// Tests for MONETcommon.F_WakeShakeWindow, the latched window in which the brake may stay open for the Wake&Shake (#151).
FUNCTION_BLOCK F_WakeShakeWindow_Tests EXTENDS TcUnit.FB_TestSuite
VAR
END_VAR

Sets_On_Exempt_Error();
Stays_Set_Without_Condition();
Not_Set_Stays_Not_Set();
Clear_Wins_Over_Set();
Timeout_Closes();
Park_Closes();
Covers_Not_Open_Closes();
Power_On_Closes();
Estop_Closes();
Other_Hw_Error_Closes();

// The #113 exemption opens the window.
METHOD PRIVATE Sets_On_Exempt_Error
VAR
	bWindow	: BOOL;
	sReason	: STRING(24);
END_VAR
TEST('Sets_On_Exempt_Error');
bWindow := MONETcommon.F_WakeShakeWindow(bWindow := FALSE, bSet := TRUE, bTimeout := FALSE, bParkActive := FALSE, bCoversOpen := TRUE, bPowerOnStart := FALSE, bEstop := FALSE, bOtherHwError := FALSE, sEndReason => sReason);
AssertTrue(Condition := bWindow, Message := 'window open');
AssertEquals_STRING(Expected := '', Actual := sReason, Message := 'no end reason');
TEST_FINISHED();
END_METHOD

// The exemption is gone after one scan; the window stays (the reason for the latch).
METHOD PRIVATE Stays_Set_Without_Condition
VAR
	bWindow	: BOOL;
	sReason	: STRING(24);
END_VAR
TEST('Stays_Set_Without_Condition');
bWindow := MONETcommon.F_WakeShakeWindow(bWindow := TRUE, bSet := FALSE, bTimeout := FALSE, bParkActive := FALSE, bCoversOpen := TRUE, bPowerOnStart := FALSE, bEstop := FALSE, bOtherHwError := FALSE, sEndReason => sReason);
AssertTrue(Condition := bWindow, Message := 'window stays open');
TEST_FINISHED();
END_METHOD

// No exemption, no window.
METHOD PRIVATE Not_Set_Stays_Not_Set
VAR
	bWindow	: BOOL;
	sReason	: STRING(24);
END_VAR
TEST('Not_Set_Stays_Not_Set');
bWindow := MONETcommon.F_WakeShakeWindow(bWindow := FALSE, bSet := FALSE, bTimeout := FALSE, bParkActive := FALSE, bCoversOpen := TRUE, bPowerOnStart := FALSE, bEstop := FALSE, bOtherHwError := FALSE, sEndReason => sReason);
AssertFalse(Condition := bWindow, Message := 'no window');
TEST_FINISHED();
END_METHOD

// Set and cleared in the same scan: not open, and no end reason (it never was open).
METHOD PRIVATE Clear_Wins_Over_Set
VAR
	bWindow	: BOOL;
	sReason	: STRING(24);
END_VAR
TEST('Clear_Wins_Over_Set');
bWindow := MONETcommon.F_WakeShakeWindow(bWindow := FALSE, bSet := TRUE, bTimeout := FALSE, bParkActive := FALSE, bCoversOpen := TRUE, bPowerOnStart := FALSE, bEstop := TRUE, bOtherHwError := FALSE, sEndReason => sReason);
AssertFalse(Condition := bWindow, Message := 'closed');
AssertEquals_STRING(Expected := '', Actual := sReason, Message := 'no reason');
TEST_FINISHED();
END_METHOD

// Window timer elapsed.
METHOD PRIVATE Timeout_Closes
VAR
	bWindow	: BOOL;
	sReason	: STRING(24);
END_VAR
TEST('Timeout_Closes');
bWindow := MONETcommon.F_WakeShakeWindow(bWindow := TRUE, bSet := FALSE, bTimeout := TRUE, bParkActive := FALSE, bCoversOpen := TRUE, bPowerOnStart := FALSE, bEstop := FALSE, bOtherHwError := FALSE, sEndReason => sReason);
AssertFalse(Condition := bWindow, Message := 'window closed');
AssertEquals_STRING(Expected := 'timeout', Actual := sReason, Message := 'reason');
TEST_FINISHED();
END_METHOD

// A park is requested, running or done.
METHOD PRIVATE Park_Closes
VAR
	bWindow	: BOOL;
	sReason	: STRING(24);
END_VAR
TEST('Park_Closes');
bWindow := MONETcommon.F_WakeShakeWindow(bWindow := TRUE, bSet := FALSE, bTimeout := FALSE, bParkActive := TRUE, bCoversOpen := TRUE, bPowerOnStart := FALSE, bEstop := FALSE, bOtherHwError := FALSE, sEndReason => sReason);
AssertFalse(Condition := bWindow, Message := 'window closed');
AssertEquals_STRING(Expected := 'park', Actual := sReason, Message := 'reason');
TEST_FINISHED();
END_METHOD

// The covers are not open any more.
METHOD PRIVATE Covers_Not_Open_Closes
VAR
	bWindow	: BOOL;
	sReason	: STRING(24);
END_VAR
TEST('Covers_Not_Open_Closes');
bWindow := MONETcommon.F_WakeShakeWindow(bWindow := TRUE, bSet := FALSE, bTimeout := FALSE, bParkActive := FALSE, bCoversOpen := FALSE, bPowerOnStart := FALSE, bEstop := FALSE, bOtherHwError := FALSE, sEndReason => sReason);
AssertFalse(Condition := bWindow, Message := 'window closed');
AssertEquals_STRING(Expected := 'covers not open', Actual := sReason, Message := 'reason');
TEST_FINISHED();
END_METHOD

// A new power-on enables the elevation.
METHOD PRIVATE Power_On_Closes
VAR
	bWindow	: BOOL;
	sReason	: STRING(24);
END_VAR
TEST('Power_On_Closes');
bWindow := MONETcommon.F_WakeShakeWindow(bWindow := TRUE, bSet := FALSE, bTimeout := FALSE, bParkActive := FALSE, bCoversOpen := TRUE, bPowerOnStart := TRUE, bEstop := FALSE, bOtherHwError := FALSE, sEndReason => sReason);
AssertFalse(Condition := bWindow, Message := 'window closed');
AssertEquals_STRING(Expected := 'power-on', Actual := sReason, Message := 'reason');
TEST_FINISHED();
END_METHOD

// E-stop.
METHOD PRIVATE Estop_Closes
VAR
	bWindow	: BOOL;
	sReason	: STRING(24);
END_VAR
TEST('Estop_Closes');
bWindow := MONETcommon.F_WakeShakeWindow(bWindow := TRUE, bSet := FALSE, bTimeout := FALSE, bParkActive := FALSE, bCoversOpen := TRUE, bPowerOnStart := FALSE, bEstop := TRUE, bOtherHwError := FALSE, sEndReason => sReason);
AssertFalse(Condition := bWindow, Message := 'window closed');
AssertEquals_STRING(Expected := 'E-stop', Actual := sReason, Message := 'reason');
TEST_FINISHED();
END_METHOD

// Focus or derotator error.
METHOD PRIVATE Other_Hw_Error_Closes
VAR
	bWindow	: BOOL;
	sReason	: STRING(24);
END_VAR
TEST('Other_Hw_Error_Closes');
bWindow := MONETcommon.F_WakeShakeWindow(bWindow := TRUE, bSet := FALSE, bTimeout := FALSE, bParkActive := FALSE, bCoversOpen := TRUE, bPowerOnStart := FALSE, bEstop := FALSE, bOtherHwError := TRUE, sEndReason => sReason);
AssertFalse(Condition := bWindow, Message := 'window closed');
AssertEquals_STRING(Expected := 'focus/derotator error', Actual := sReason, Message := 'reason');
TEST_FINISHED();
END_METHOD

END_FUNCTION_BLOCK

(* stored: Version 1.1.0.1, ProductVersion 3.1.4024.15
   POU F_WakeShakeWindow_Tests: Id {365afcba-9976-43a0-b37b-22b72c50967f}, SpecialFunc None
   Method Sets_On_Exempt_Error: Id {3439bf1a-0345-4420-88a1-fdbd0de5eb7b}
   Method Stays_Set_Without_Condition: Id {3c26585b-2306-43d8-8add-422688d4f568}
   Method Not_Set_Stays_Not_Set: Id {72ca0856-d219-44b0-93e0-4150c6ed9e9f}
   Method Clear_Wins_Over_Set: Id {2a60a101-e590-487f-a56f-42d655a0d487}
   Method Timeout_Closes: Id {7bf0f4b7-0611-4a2f-816d-bdca26f6d4d7}
   Method Park_Closes: Id {66d89e64-c0e1-45f8-8420-dc79337b6856}
   Method Covers_Not_Open_Closes: Id {0b32e7ae-2341-4232-95f8-79c68a7b7d1e}
   Method Power_On_Closes: Id {6d2ae647-6bd8-48f8-8146-77ad3e83c70c}
   Method Estop_Closes: Id {7ec98f05-e44b-4a85-a68d-1a61f0b35381}
   Method Other_Hw_Error_Closes: Id {66b42fc4-8815-4cd1-ae7d-96a5822ac11b} *)
